(* IEC 61131-3 sources: codesys-to-astra/corpus/s7-chain/src/POUs/S7Compat/FB_S7Tp, 2 files *)

(* ---- FB_S7Tp.decl.st ---- *)
// Назначение: импульсный таймер с интерфейсом TP (IN, PT, Q, ET) для кода, сконвертированного s7conv
//             из S7 TP_TIME/TP с --timers s7compat. Семантика МЭК 61131-3 и S7: фронт IN вне импульса
//             запускает импульс Q длительностью PT; фронты во время импульса его не продлевают; ET
//             растёт до PT во время импульса, после импульса остаётся PT, пока IN = TRUE, и
//             сбрасывается в 0 при IN = FALSE. Время — F_S7Now(): в работе TIME(), как у Standard.TP,
//             в тестах — моделируемые часы GVL_S7Clock. Совпадение со Standard.TP в реальном времени —
//             тест FB_S7Tp_Test.MatchesStandardInRealTime.
// Автор:      kr0nsch
// Версия:     0.1.0
// Документ:   docs/MAPPING.md, раздел «Функциональные блоки инструкций»; docs/methodology.md
FUNCTION_BLOCK FB_S7Tp
VAR_INPUT
    IN : BOOL;          // lint:allow STL007 интерфейс TP: имя входа как у Standard.TP
    PT : TIME;          // lint:allow STL007 интерфейс TP: длительность импульса
END_VAR
VAR_OUTPUT
    Q : BOOL;           // lint:allow STL007 интерфейс TP: импульс
    ET : TIME;          // lint:allow STL007 интерфейс TP: прошедшее время импульса
END_VAR
VAR
    xInPrev : BOOL;     // IN на прошлом вызове (FALSE до первого вызова)
    tNow : TIME;        // время этого вызова (F_S7Now читается один раз)
    tStart : TIME;      // начало импульса
    tElapsed : TIME;    // прошло с tStart
END_VAR

(* ---- FB_S7Tp.impl.st ---- *)
tNow := F_S7Now();
// фронт IN вне импульса: начало импульса
IF IN AND NOT xInPrev AND NOT Q THEN
    tStart := tNow;
    Q := TRUE;
END_IF

IF Q THEN
    tElapsed := tNow - tStart;
    IF tElapsed >= PT THEN
        Q := FALSE;
        ET := PT;
    ELSE
        ET := tElapsed;
    END_IF
END_IF

// импульса нет и IN = FALSE: ET сбрасывается (после импульса при IN = TRUE ET = PT)
IF NOT IN AND NOT Q THEN
    ET := T#0MS;
END_IF
xInPrev := IN;
